TYPE (* The fixed type hash *)
  (* Standard: 61499-1; Description: Copyright (c) 2026 Osoft e.U. This program and the accompanying materials are made available under the terms of the Eclipse Public License 2.0 which is available at https://www.eclipse.org/legal/epl-2.0/ SPDX-License-Identifier: EPL-2.0 *)
  (* Version 1.0, 2026-11-19, Michael Oberlehner, initial API and implementation and/or initial documentation *)
  PACKAGE eclipse4diac::core;
  TypeHash : STRING := ''; (* The fixed type hash *)
END_TYPE
